(* PLC project motor, tcpethernet motor 1 *)
(* stored: creationDateTime 2026-10-28T09:00:00, modificationDateTime 2026-10-28T09:00:00 *)

PROGRAM motor
  VAR
    Start AT %IX0.0 : BOOL;
    Stop AT %IX0.1 : BOOL;
    Lamp AT %QX0.0 : BOOL;
  END_VAR
  VAR
    Run : BOOL;
    Fan : BOOL;
    delay : TON;
  END_VAR

(* LD diagram, written out as Structured Text *)
Run := (Start OR Run) AND NOT Stop;
Lamp := (Start OR Run) AND NOT Stop;
delay(IN := Run, PT := T#2s);
Fan := delay.Q;
END_PROGRAM

CONFIGURATION config
  RESOURCE resource1 ON PLC
    TASK main(INTERVAL := T#10ms, PRIORITY := 0);
    PROGRAM instance0 WITH main : motor;
  END_RESOURCE
END_CONFIGURATION
